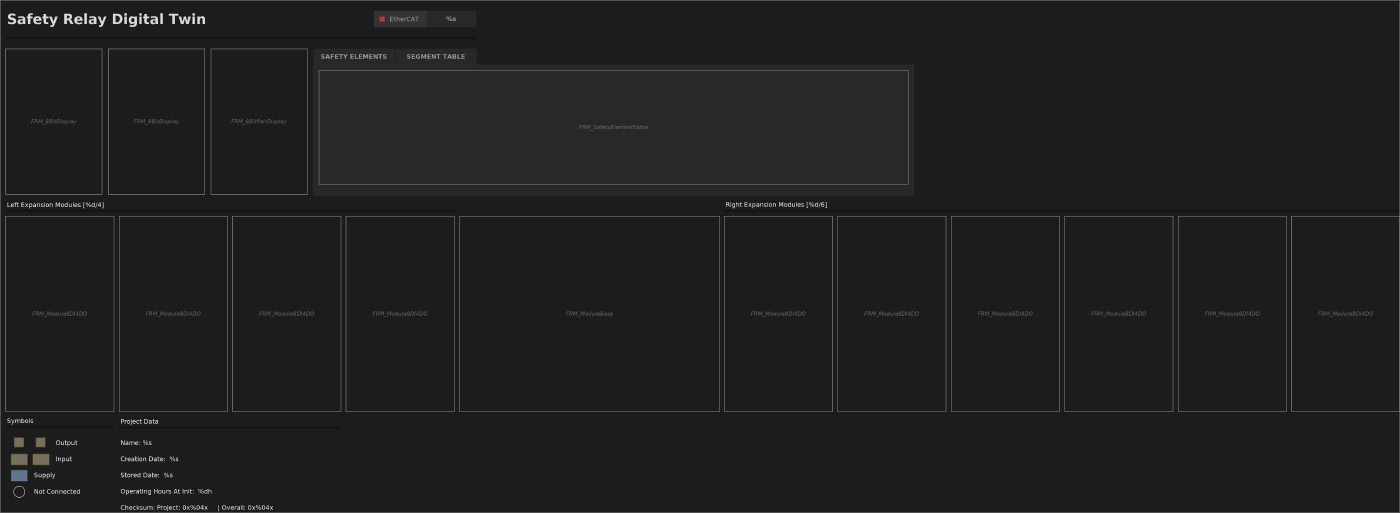
VISUALIZATION Safety  // 2591x950
VAR
    nTabIndex: USINT := 0;
   bUnused: BOOL := FALSE;
END_VAR
    Line (10,70) (882,70)
    Label (10,10 421x51), "Safety Relay Digital Twin"
    Frame (200,90 179x270)
        shows FRM_8BitDisplay(sName := 'O Bits', sBit0 := 'Heartbeat', sBit1 := 'Ack. Required', sBit2 := 'Message', sBit3 := 'Warning', sBit4 := 'Message', sBit5 := 'E-Stop OK', sBit6 := 'Remote', sBit7 := '-', bBit0 := Motion_Safety.stSafety.stIn.stMCCStatus.bHeartbeat, bBit1 := Motion_Safety.stSafety.stIn.stMCCStatus.bAcknowledgeRequired, bBit2 := Motion_Safety.stSafety.stIn.stMCCStatus.bFault, bBit3 := Motion_Safety.stSafety.stIn.stMCCStatus.bWarning, bBit4 := Motion_Safety.stSafety.stIn.stMCCStatus.bMessage, bBit5 := Motion_Safety.stSafety.stIn.stMCCStatus.bEStopOK, bBit6 := Motion_Safety.stSafety.stIn.stMCCStatus.bRemote, bBit7 := bUnused)
    Frame (10,90 179x270)
        shows FRM_8BitDisplay(sName := 'I Bits', sBit0 := 'Heartbeat', sBit1 := 'PLC OK', sBit2 := 'Error Ack.', sBit3 := '-', sBit4 := '-', sBit5 := '-', sBit6 := '-', sBit7 := '-', bBit0 := Motion_Safety.stSafety.stOut.stMCCStatus.bHeartbeat, bBit1 := Motion_Safety.stSafety.stOut.stMCCStatus.bPLC_OK, bBit2 := Motion_Safety.stSafety.stOut.stMCCStatus.bErrorAcknowledge, bBit3 := bUnused, bBit4 := bUnused, bBit5 := bUnused, bBit6 := bUnused, bBit7 := bUnused)
    Frame (390,90 179x270)
        shows FRM_8BitPairDisplay(bBit0_1 := Motion_Safety.stSafety.stIn.stMCCAppSpecific.abData[1], bBit1_1 := Motion_Safety.stSafety.stIn.stMCCAppSpecific.abData[2], bBit2_1 := Motion_Safety.stSafety.stIn.stMCCAppSpecific.abData[3], bBit3_1 := Motion_Safety.stSafety.stIn.stMCCAppSpecific.abData[4], bBit4_1 := Motion_Safety.stSafety.stIn.stMCCAppSpecific.abData[5], bBit5_1 := Motion_Safety.stSafety.stIn.stMCCAppSpecific.abData[6], bBit6_1 := Motion_Safety.stSafety.stIn.stMCCAppSpecific.abData[7], bBit7_1 := Motion_Safety.stSafety.stIn.stMCCAppSpecific.abData[8], bBit0_2 := Motion_Safety.stSafety.stIn.stMCCAppSpecific.abValid[1], bBit1_2 := Motion_Safety.stSafety.stIn.stMCCAppSpecific.abValid[2], bBit2_2 := Motion_Safety.stSafety.stIn.stMCCAppSpecific.abValid[3], bBit3_2 := Motion_Safety.stSafety.stIn.stMCCAppSpecific.abValid[4], bBit4_2 := Motion_Safety.stSafety.stIn.stMCCAppSpecific.abValid[5], bBit5_2 := Motion_Safety.stSafety.stIn.stMCCAppSpecific.abValid[6], bBit6_2 := Motion_Safety.stSafety.stIn.stMCCAppSpecific.abValid[7], bBit7_2 := Motion_Safety.stSafety.stIn.stMCCAppSpecific.abValid[8], sName := 'APPLICATION', sBitPair0 := 'App 1', sBitPair1 := 'App 2', sBitPair2 := 'App 3', sBitPair3 := 'App 4', sBitPair4 := 'App 5', sBitPair5 := 'App 6', sBitPair6 := 'App 7', sBitPair7 := 'App 8')
    Ellipse (25,900 21x21)
    Label (100,810 51x20), "Output"
    Label (100,840 51x20), "Input"
    Label (60,870 51x20), "Supply"
    Label (60,900 101x21), "Not Connected"
    Rectangle (20,840 31x21)
    Rectangle (20,870 31x21)
    Rectangle (26,810 18x18), angle 45
    Rectangle (60,840 31x21), colour toggle: TRUE
    Rectangle (66,810 18x18), angle 45, colour toggle: TRUE
    Rectangle (580,120 1111x241)
    Frame (590,130 1091x211)
        shows FRM_SafetyElementTable(nFunctionCount := GVL_APP.nNUM_OF_SAFE_FUNCTIONS, nInputCount := GVL_APP.nNUM_OF_SAFE_INPUTS, nOutputCount := GVL_APP.nNUM_OF_SAFE_OUTPUTS)
        shows FRM_SegmentTable(nRequestTableNo := Motion_Safety.fbMotionSafety.stPNOZEtherCATOut.nTableNumber, nRequestSegmentNo := Motion_Safety.fbMotionSafety.stPNOZEtherCATOut.nSegmentNumber, nResponseTableNo := Motion_Safety.fbMotionSafety.stPNOZEtherCATIn.nTableNumber, nResponseSegmentNo := Motion_Safety.fbMotionSafety.stPNOZEtherCATIn.nSegmentNumber, aSegmentBytes := Motion_Safety.fbMotionSafety.stPNOZEtherCATIn.anSegmentByte)
    Rectangle (580,90 150x30), "SAFETY ELEMENTS", colour toggle: nTabIndex = 0
        OnMouseUp: execute { nTabIndex := 0; }
        OnMouseUp: FrameSelectionChange Selection=SelectedFrame=2ac8e0da-98ce-4fdd-a785-8dd91d41c461, GlobSel=AssignType=Directly, SelType=Locally
    Rectangle (732,90 150x30), "SEGMENT TABLE", colour toggle: nTabIndex = 1
        OnMouseUp: execute { nTabIndex := 1; }
        OnMouseUp: FrameSelectionChange Selection=SelectedFrame=2ac8e0da-98ce-4fdd-a785-8dd91d41c461, Selection=1, GlobSel=AssignType=Directly, SelType=Locally
    Rectangle (692,20 99x30)
    Rectangle (702,30 10x10), colour toggle: Motion_Safety.stSafety.stIn.stPNOZCommDiag.nEtherCATState > 4
    Frame (1340,400 201x362), invisible if: GVL_APP.nNUM_OF_EXPANSION_RIGHT < 1, frame switch variable: Motion_Safety.stSafety.stIn.astExpansionModuleRightData[1].eDeviceType
        shows FRM_Module8DI4DO(stModuleData := Motion_Safety.stSafety.stIn.astExpansionModuleRightData[1], nIndex := 1)
        shows FRM_Module4DI4DOR(stModuleData := Motion_Safety.stSafety.stIn.astExpansionModuleRightData[1], nIndex := 1)
        p3528305787: -210 * ( GVL_APP.nMAX_EXPANSION_MODULE_LEFT - GVL_APP.nNUM_OF_EXPANSION_LEFT)
    Frame (1550,400 201x362), invisible if: GVL_APP.nNUM_OF_EXPANSION_RIGHT < 2, frame switch variable: Motion_Safety.stSafety.stIn.astExpansionModuleRightData[2].eDeviceType
        shows FRM_Module8DI4DO(stModuleData := Motion_Safety.stSafety.stIn.astExpansionModuleRightData[2], nIndex := 2)
        shows FRM_Module4DI4DOR(stModuleData := Motion_Safety.stSafety.stIn.astExpansionModuleRightData[2], nIndex := 2)
        p3528305787: -210 * ( GVL_APP.nMAX_EXPANSION_MODULE_LEFT - GVL_APP.nNUM_OF_EXPANSION_LEFT)
    Frame (1760,400 201x362), invisible if: GVL_APP.nNUM_OF_EXPANSION_RIGHT < 3, frame switch variable: Motion_Safety.stSafety.stIn.astExpansionModuleRightData[3].eDeviceType
        shows FRM_Module8DI4DO(stModuleData := Motion_Safety.stSafety.stIn.astExpansionModuleRightData[3], nIndex := 3)
        shows FRM_Module4DI4DOR(stModuleData := Motion_Safety.stSafety.stIn.astExpansionModuleRightData[3], nIndex := 3)
        p3528305787: -210 * ( GVL_APP.nMAX_EXPANSION_MODULE_LEFT - GVL_APP.nNUM_OF_EXPANSION_LEFT)
    Frame (1970,400 201x362), invisible if: GVL_APP.nNUM_OF_EXPANSION_RIGHT < 4, frame switch variable: Motion_Safety.stSafety.stIn.astExpansionModuleRightData[4].eDeviceType
        shows FRM_Module8DI4DO(stModuleData := Motion_Safety.stSafety.stIn.astExpansionModuleRightData[4], nIndex := 4)
        shows FRM_Module4DI4DOR(stModuleData := Motion_Safety.stSafety.stIn.astExpansionModuleRightData[4], nIndex := 4)
        p3528305787: -210 * ( GVL_APP.nMAX_EXPANSION_MODULE_LEFT - GVL_APP.nNUM_OF_EXPANSION_LEFT)
    Label (718,20 61x31), "EtherCAT"
    Rectangle (790,20 91x30), "%s", text variable: Motion_Safety.fbMotionSafety.sEtherCATState
    Frame (2180,400 201x362), invisible if: GVL_APP.nNUM_OF_EXPANSION_RIGHT < 5, frame switch variable: Motion_Safety.stSafety.stIn.astExpansionModuleRightData[5].eDeviceType
        shows FRM_Module8DI4DO(stModuleData := Motion_Safety.stSafety.stIn.astExpansionModuleRightData[5], nIndex := 5)
        shows FRM_Module4DI4DOR(stModuleData := Motion_Safety.stSafety.stIn.astExpansionModuleRightData[5], nIndex := 5)
        p3528305787: -210 * ( GVL_APP.nMAX_EXPANSION_MODULE_LEFT - GVL_APP.nNUM_OF_EXPANSION_LEFT)
    Frame (2390,400 201x362), invisible if: GVL_APP.nNUM_OF_EXPANSION_RIGHT < 6, frame switch variable: Motion_Safety.stSafety.stIn.astExpansionModuleRightData[6].eDeviceType
        shows FRM_Module8DI4DO(stModuleData := Motion_Safety.stSafety.stIn.astExpansionModuleRightData[6], nIndex := 6)
        shows FRM_Module4DI4DOR(stModuleData := Motion_Safety.stSafety.stIn.astExpansionModuleRightData[6], nIndex := 6)
        p3528305787: -210 * ( GVL_APP.nMAX_EXPANSION_MODULE_LEFT - GVL_APP.nNUM_OF_EXPANSION_LEFT)
    Frame (850,400 482x362)
        shows FRM_ModuleBase(stFieldbusData := Motion_Safety.stSafety.stIn.stFieldbusData, stBaseModuleData := Motion_Safety.stSafety.stIn.stBaseModuleData)
        p3528305787: -210 * ( GVL_APP.nMAX_EXPANSION_MODULE_LEFT - GVL_APP.nNUM_OF_EXPANSION_LEFT)
    Frame (10,400 201x362), invisible if: GVL_APP.nNUM_OF_EXPANSION_LEFT < 4, frame switch variable: Motion_Safety.stSafety.stIn.astExpansionModuleLeftData[4].eDeviceType
        shows FRM_Module8DI4DO(stModuleData := Motion_Safety.stSafety.stIn.astExpansionModuleLeftData[4], nIndex := 4)
        shows FRM_Module4DI4DOR(stModuleData := Motion_Safety.stSafety.stIn.astExpansionModuleLeftData[4], nIndex := 4)
    Frame (220,400 201x362), invisible if: GVL_APP.nNUM_OF_EXPANSION_LEFT < 3, frame switch variable: Motion_Safety.stSafety.stIn.astExpansionModuleLeftData[3].eDeviceType
        shows FRM_Module8DI4DO(stModuleData := Motion_Safety.stSafety.stIn.astExpansionModuleLeftData[3], nIndex := 3)
        shows FRM_Module4DI4DOR(stModuleData := Motion_Safety.stSafety.stIn.astExpansionModuleLeftData[3], nIndex := 3)
        p3528305787: -210 * ( GVL_APP.nMAX_EXPANSION_MODULE_LEFT - GVL_APP.nNUM_OF_EXPANSION_LEFT)
    Frame (430,400 201x362), invisible if: GVL_APP.nNUM_OF_EXPANSION_LEFT < 2, frame switch variable: Motion_Safety.stSafety.stIn.astExpansionModuleLeftData[2].eDeviceType
        shows FRM_Module8DI4DO(stModuleData := Motion_Safety.stSafety.stIn.astExpansionModuleLeftData[2], nIndex := 2)
        shows FRM_Module4DI4DOR(stModuleData := Motion_Safety.stSafety.stIn.astExpansionModuleLeftData[2], nIndex := 2)
        p3528305787: -210 * ( GVL_APP.nMAX_EXPANSION_MODULE_LEFT - GVL_APP.nNUM_OF_EXPANSION_LEFT)
    Frame (640,400 201x362), invisible if: GVL_APP.nNUM_OF_EXPANSION_LEFT < 1, frame switch variable: Motion_Safety.stSafety.stIn.astExpansionModuleLeftData[1].eDeviceType
        shows FRM_Module8DI4DO(stModuleData := Motion_Safety.stSafety.stIn.astExpansionModuleLeftData[1], nIndex := 1)
        shows FRM_Module4DI4DOR(stModuleData := Motion_Safety.stSafety.stIn.astExpansionModuleLeftData[1], nIndex := 1)
        p3528305787: -210 * ( GVL_APP.nMAX_EXPANSION_MODULE_LEFT - GVL_APP.nNUM_OF_EXPANSION_LEFT)
    Line (10,790) (210,790)
    Line (10,390) (840,390), invisible if: GVL_APP.nNUM_OF_EXPANSION_LEFT < 1
        p874137650: -210 * ( GVL_APP.nMAX_EXPANSION_MODULE_LEFT - GVL_APP.nNUM_OF_EXPANSION_LEFT)
    Line (1340,390) (2590,390), invisible if: GVL_APP.nNUM_OF_EXPANSION_RIGHT < 1
        p3528305787: -210 * ( GVL_APP.nMAX_EXPANSION_MODULE_LEFT - GVL_APP.nNUM_OF_EXPANSION_LEFT)
        p874137650: -210 * ( GVL_APP.nMAX_EXPANSION_MODULE_LEFT - GVL_APP.nNUM_OF_EXPANSION_LEFT) - 210 * ( GVL_APP.nMAX_EXPANSION_MODULE_RIGHT - GVL_APP.nNUM_OF_EXPANSION_RIGHT)
    Rectangle (10,369 251x21), "Left Expansion Modules [%d/4]", text variable: GVL_APP.nNUM_OF_EXPANSION_LEFT, invisible if: GVL_APP.nNUM_OF_EXPANSION_LEFT < 1
    Rectangle (1340,369 251x20), "Right Expansion Modules [%d/6]", text variable: GVL_APP.nNUM_OF_EXPANSION_RIGHT, invisible if: GVL_APP.nNUM_OF_EXPANSION_RIGHT < 1
        p3528305787: -210 * ( GVL_APP.nMAX_EXPANSION_MODULE_LEFT - GVL_APP.nNUM_OF_EXPANSION_LEFT)
    Label (10,769 91x21), "Symbols"
    Line (220,791) (630,791)
    Label (220,770 91x21), "Project Data"
    Textfield (220,810 411x20), "Name: %s", text variable: Motion_Safety.fbMotionSafety.fbPNOZData.stData.wsProjectName
    Textfield (220,840 321x20), "Creation Date: %s", text variable: Motion_Safety.fbMotionSafety.fbPNOZData.stData.sCreationDate
    Textfield (220,930 181x20), "Checksum: Project: 0x%04x", text variable: Motion_Safety.fbMotionSafety.fbPNOZData.stData.nProjectChecksum
    Textfield (400,930 231x20), "| Overall: 0x%04x", text variable: Motion_Safety.fbMotionSafety.fbPNOZData.stData.nOverallChecksum
    Textfield (220,870 321x20), "Stored Date: %s", text variable: Motion_Safety.fbMotionSafety.fbPNOZData.stData.sStoredDate
    Textfield (220,900 411x20), "Operating Hours At Init: %dh", text variable: Motion_Safety.fbMotionSafety.fbPNOZData.stData.nOperatingHoursAtInit
END_VISUALIZATION

(* stored: Version 1.1.0.1
   Visu Safety: Id {0e6e1981-dea2-07f9-2a3d-84624e740091} *)
